(* IEC 61131-3 sources: rusty/tests/lit/single/type_promotion/bit_string/unary_minus, 2 files *)

(* ---- byte_word_operand.st ---- *)
// RUN: %COMPILE %s && %RUN | %CHECK %s
// The negation of a BYTE or WORD is computed in DINT, so a value from the signed midpoint on gives the negative value.
FUNCTION main : DINT
    VAR
        b : BYTE := 16#FF;
        b200 : BYTE := 16#C8;
        w : WORD := 16#FFFF;
        w40000 : WORD := 16#9C40;
        r : LINT;
    END_VAR

    r := -b;
    printf('-BYTE 16#FF = %lld$N', r);                      // CHECK: -BYTE 16#FF = -255
    r := -b200;
    printf('-BYTE 16#C8 = %lld$N', r);                      // CHECK-NEXT: -BYTE 16#C8 = -200
    r := -w;
    printf('-WORD 16#FFFF = %lld$N', r);                    // CHECK-NEXT: -WORD 16#FFFF = -65535
    r := -w40000;
    printf('-WORD 16#9C40 = %lld$N', r);                    // CHECK-NEXT: -WORD 16#9C40 = -40000
    printf('-BYTE 16#FF < 0 = %d$N', -b < 0);               // CHECK-NEXT: -BYTE 16#FF < 0 = 1
END_FUNCTION

(* ---- dword_operand.st ---- *)
// RUN: %COMPILE %s && %RUN | %CHECK %s
// The negation of a DWORD is LINT, so a value from 2^31 on gives the negative value.
FUNCTION main : DINT
    VAR
        dw : DWORD := 16#FFFF_FFFF;
        dw3e9 : DWORD := 16#B2D0_5E00;
        r : LINT;
    END_VAR

    r := -dw;
    printf('-DWORD 16#FFFF_FFFF = %lld$N', r);              // CHECK: -DWORD 16#FFFF_FFFF = -4294967295
    r := -dw3e9;
    printf('-DWORD 16#B2D0_5E00 = %lld$N', r);              // CHECK-NEXT: -DWORD 16#B2D0_5E00 = -3000000000
END_FUNCTION
